// LS Electric XG5000 project: 신호등
// PLC LSPLC

PROGRAM NewProgram (task: 스캔 프로그램)

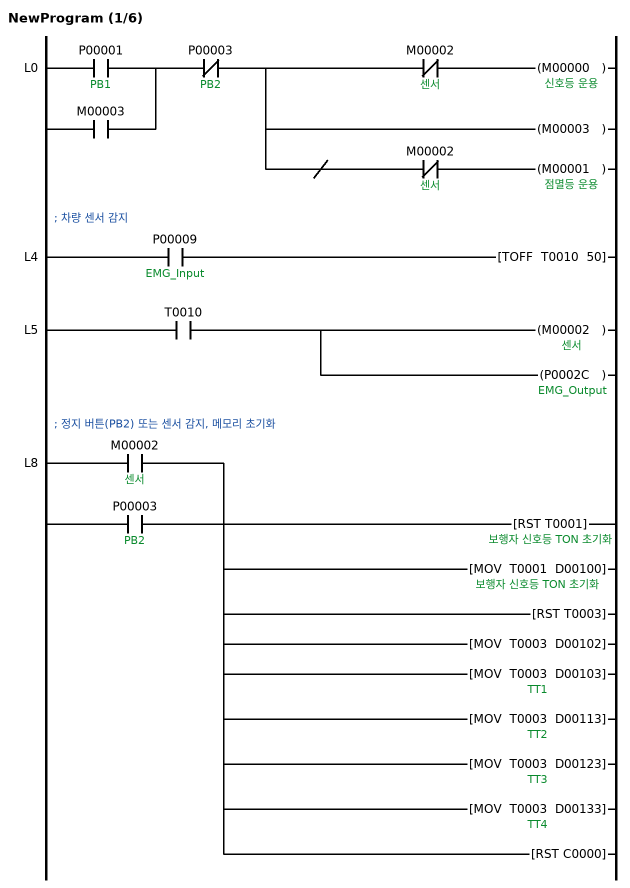
; L0
LOAD      P00001	// PB1
OR        M00003
AND NOT   P00003	// PB2
MPUSH
AND NOT   M00002	// 센서
OUT       M00000	// 신호등 운용
MPOP
OUT       M00003
NOT
AND NOT   M00002	// 센서
OUT       M00001	// 점멸등 운용
// 차량 센서 감지
; L4
LOAD      P00009	// EMG_Input
TOFF      T0010 50
; L5
LOAD      T0010
OUT       M00002	// 센서
OUT       P0002C	// EMG_Output
// 정지 버튼(PB2) 또는 센서 감지, 메모리 초기화
; L8
LOAD      M00002	// 센서
OR        P00003	// PB2
RST       T0001	// 보행자 신호등 TON 초기화
MOV       T0001 D00100	// 보행자 신호등 TON 초기화
RST       T0003
MOV       T0003 D00102
MOV       T0003 D00103	// TT1
MOV       T0003 D00113	// TT2
MOV       T0003 D00123	// TT3
MOV       T0003 D00133	// TT4
RST       C0000

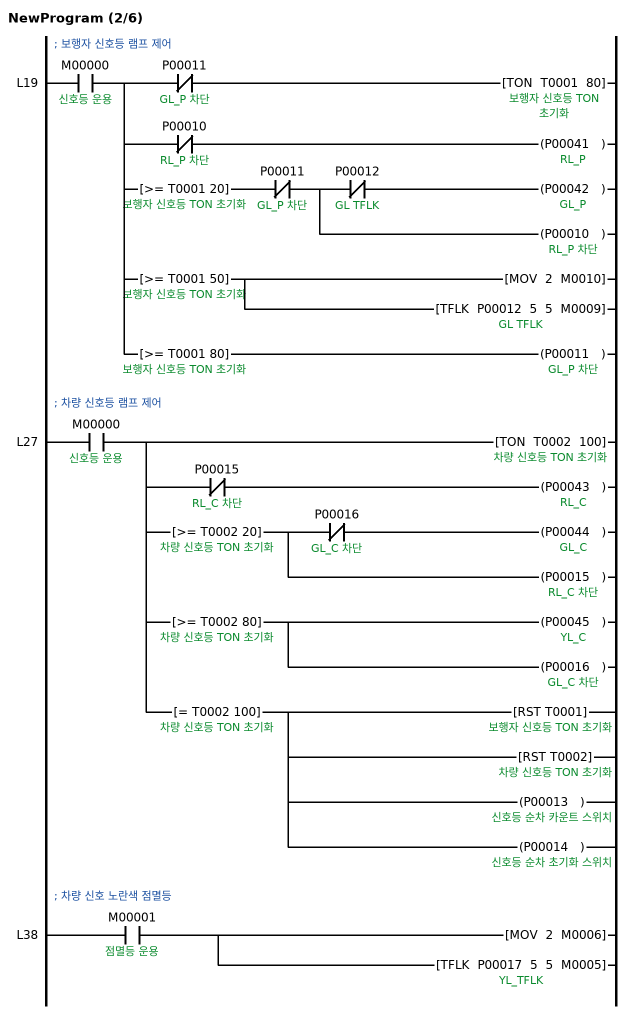
// 보행자 신호등 램프 제어
; L19
LOAD      M00000	// 신호등 운용
MPUSH
AND NOT   P00011	// GL_P 차단
TON       T0001 80	// 보행자 신호등 TON 초기화
MLOAD
AND NOT   P00010	// RL_P 차단
OUT       P00041	// RL_P
MLOAD
AND>=     T0001 20	// 보행자 신호등 TON 초기화
AND NOT   P00011	// GL_P 차단
MPUSH
AND NOT   P00012	// GL TFLK
OUT       P00042	// GL_P
MPOP
OUT       P00010	// RL_P 차단
MLOAD
AND>=     T0001 50	// 보행자 신호등 TON 초기화
MOV       2 M0010
TFLK      P00012 5 5 M0009	// GL TFLK
MPOP
AND>=     T0001 80	// 보행자 신호등 TON 초기화
OUT       P00011	// GL_P 차단
// 차량 신호등 램프 제어
; L27
LOAD      M00000	// 신호등 운용
TON       T0002 100	// 차량 신호등 TON 초기화
MPUSH
AND NOT   P00015	// RL_C 차단
OUT       P00043	// RL_C
MLOAD
AND>=     T0002 20	// 차량 신호등 TON 초기화
MPUSH
AND NOT   P00016	// GL_C 차단
OUT       P00044	// GL_C
MPOP
OUT       P00015	// RL_C 차단
MLOAD
AND>=     T0002 80	// 차량 신호등 TON 초기화
OUT       P00045	// YL_C
OUT       P00016	// GL_C 차단
MPOP
AND=      T0002 100	// 차량 신호등 TON 초기화
RST       T0001	// 보행자 신호등 TON 초기화
RST       T0002	// 차량 신호등 TON 초기화
OUT       P00013	// 신호등 순차 카운트 스위치
OUT       P00014	// 신호등 순차 초기화 스위치
// 차량 신호 노란색 점멸등
; L38
LOAD      M00001	// 점멸등 운용
MOV       2 M0006
TFLK      P00017 5 5 M0005	// YL_TFLK

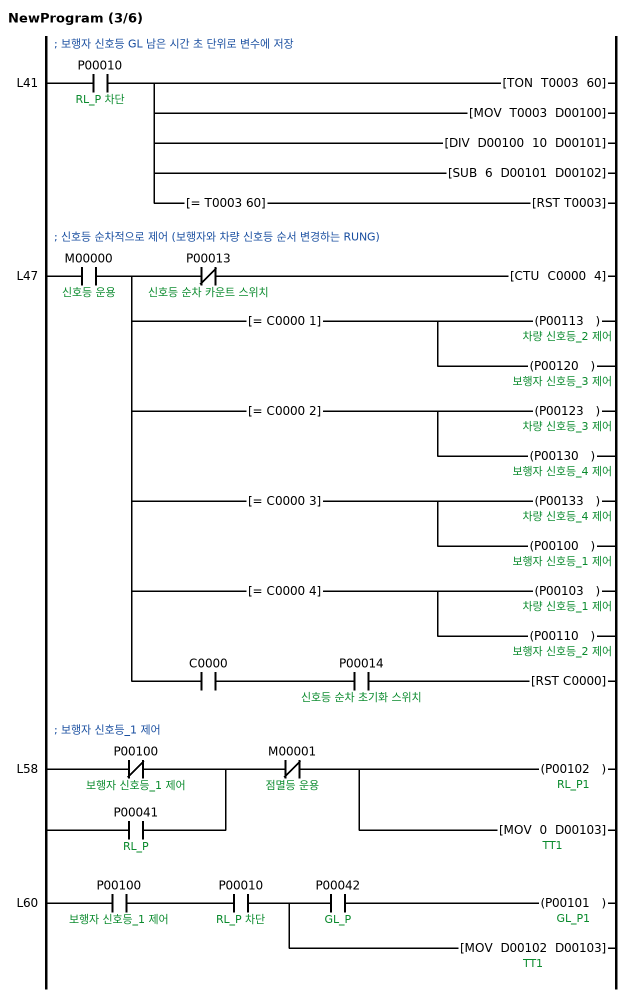
// 보행자 신호등 GL 남은 시간 초 단위로 변수에 저장
; L41
LOAD      P00010	// RL_P 차단
TON       T0003 60
MOV       T0003 D00100
DIV       D00100 10 D00101
SUB       6 D00101 D00102
AND=      T0003 60
RST       T0003
// 신호등 순차적으로 제어 (보행자와 차량 신호등 순서 변경하는 RUNG)
; L47
LOAD      M00000	// 신호등 운용
MPUSH
AND NOT   P00013	// 신호등 순차 카운트 스위치
CTU       C0000 4
MLOAD
AND=      C0000 1
OUT       P00113	// 차량 신호등_2 제어
OUT       P00120	// 보행자 신호등_3 제어
MLOAD
AND=      C0000 2
OUT       P00123	// 차량 신호등_3 제어
OUT       P00130	// 보행자 신호등_4 제어
MLOAD
AND=      C0000 3
OUT       P00133	// 차량 신호등_4 제어
OUT       P00100	// 보행자 신호등_1 제어
MLOAD
AND=      C0000 4
OUT       P00103	// 차량 신호등_1 제어
OUT       P00110	// 보행자 신호등_2 제어
MPOP
AND       C0000
AND       P00014	// 신호등 순차 초기화 스위치
RST       C0000
// 보행자 신호등_1 제어
; L58
LOAD NOT  P00100	// 보행자 신호등_1 제어
OR        P00041	// RL_P
AND NOT   M00001	// 점멸등 운용
OUT       P00102	// RL_P1
MOV       0 D00103	// TT1
; L60
LOAD      P00100	// 보행자 신호등_1 제어
AND       P00010	// RL_P 차단
MPUSH
AND       P00042	// GL_P
OUT       P00101	// GL_P1
MPOP
MOV       D00102 D00103	// TT1

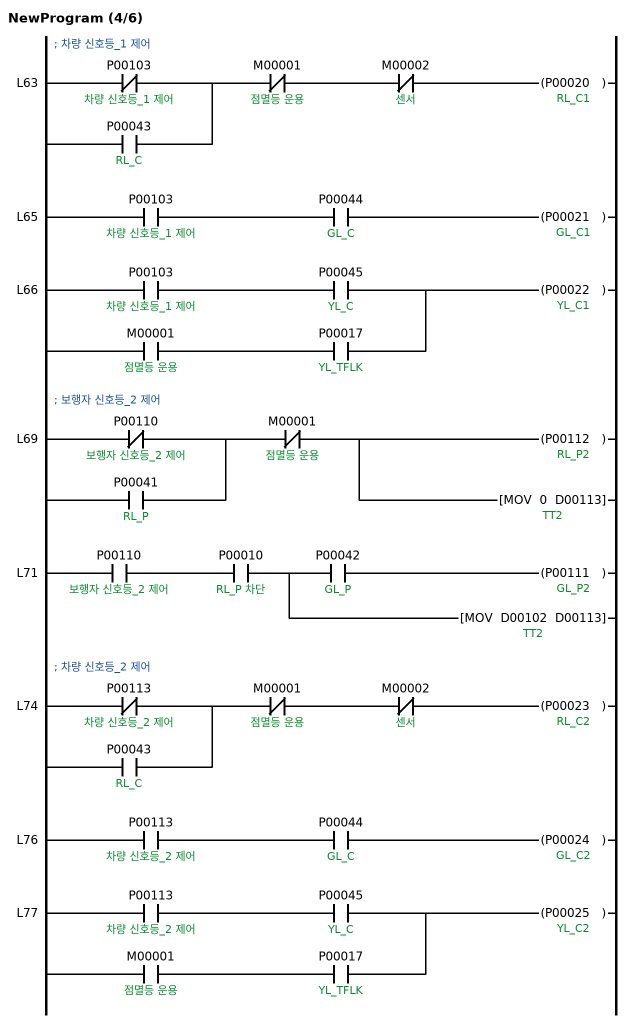
// 차량 신호등_1 제어
; L63
LOAD NOT  P00103	// 차량 신호등_1 제어
OR        P00043	// RL_C
AND NOT   M00001	// 점멸등 운용
AND NOT   M00002	// 센서
OUT       P00020	// RL_C1
; L65
LOAD      P00103	// 차량 신호등_1 제어
AND       P00044	// GL_C
OUT       P00021	// GL_C1
; L66
LOAD      P00103	// 차량 신호등_1 제어
AND       P00045	// YL_C
LOAD      M00001	// 점멸등 운용
AND       P00017	// YL_TFLK
OR LOAD
OUT       P00022	// YL_C1
// 보행자 신호등_2 제어
; L69
LOAD NOT  P00110	// 보행자 신호등_2 제어
OR        P00041	// RL_P
AND NOT   M00001	// 점멸등 운용
OUT       P00112	// RL_P2
MOV       0 D00113	// TT2
; L71
LOAD      P00110	// 보행자 신호등_2 제어
AND       P00010	// RL_P 차단
MPUSH
AND       P00042	// GL_P
OUT       P00111	// GL_P2
MPOP
MOV       D00102 D00113	// TT2
// 차량 신호등_2 제어
; L74
LOAD NOT  P00113	// 차량 신호등_2 제어
OR        P00043	// RL_C
AND NOT   M00001	// 점멸등 운용
AND NOT   M00002	// 센서
OUT       P00023	// RL_C2
; L76
LOAD      P00113	// 차량 신호등_2 제어
AND       P00044	// GL_C
OUT       P00024	// GL_C2
; L77
LOAD      P00113	// 차량 신호등_2 제어
AND       P00045	// YL_C
LOAD      M00001	// 점멸등 운용
AND       P00017	// YL_TFLK
OR LOAD
OUT       P00025	// YL_C2

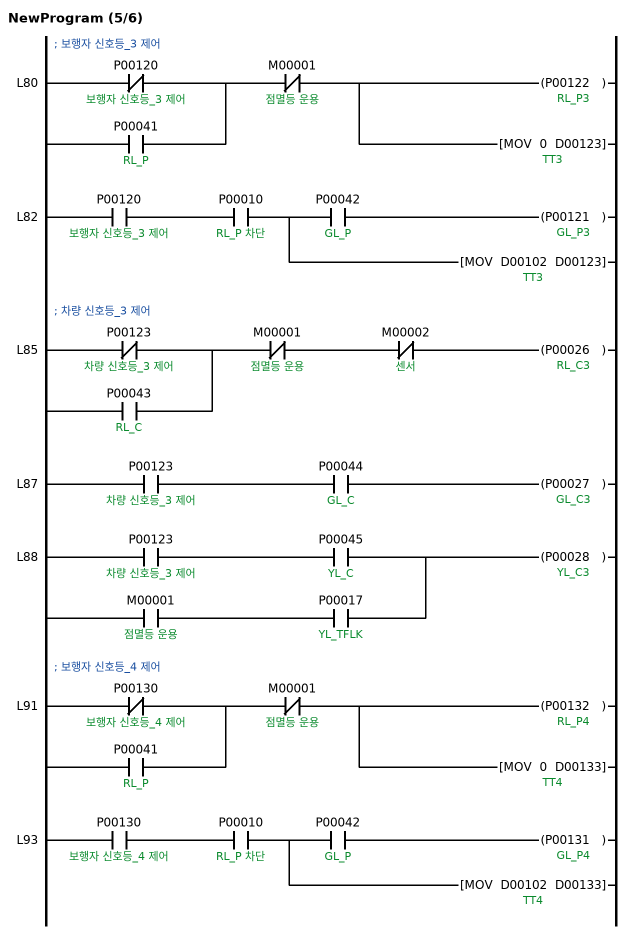
// 보행자 신호등_3 제어
; L80
LOAD NOT  P00120	// 보행자 신호등_3 제어
OR        P00041	// RL_P
AND NOT   M00001	// 점멸등 운용
OUT       P00122	// RL_P3
MOV       0 D00123	// TT3
; L82
LOAD      P00120	// 보행자 신호등_3 제어
AND       P00010	// RL_P 차단
MPUSH
AND       P00042	// GL_P
OUT       P00121	// GL_P3
MPOP
MOV       D00102 D00123	// TT3
// 차량 신호등_3 제어
; L85
LOAD NOT  P00123	// 차량 신호등_3 제어
OR        P00043	// RL_C
AND NOT   M00001	// 점멸등 운용
AND NOT   M00002	// 센서
OUT       P00026	// RL_C3
; L87
LOAD      P00123	// 차량 신호등_3 제어
AND       P00044	// GL_C
OUT       P00027	// GL_C3
; L88
LOAD      P00123	// 차량 신호등_3 제어
AND       P00045	// YL_C
LOAD      M00001	// 점멸등 운용
AND       P00017	// YL_TFLK
OR LOAD
OUT       P00028	// YL_C3
// 보행자 신호등_4 제어
; L91
LOAD NOT  P00130	// 보행자 신호등_4 제어
OR        P00041	// RL_P
AND NOT   M00001	// 점멸등 운용
OUT       P00132	// RL_P4
MOV       0 D00133	// TT4
; L93
LOAD      P00130	// 보행자 신호등_4 제어
AND       P00010	// RL_P 차단
MPUSH
AND       P00042	// GL_P
OUT       P00131	// GL_P4
MPOP
MOV       D00102 D00133	// TT4

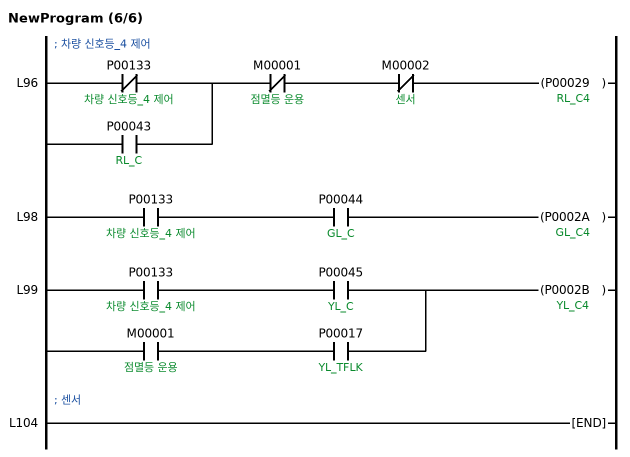
// 차량 신호등_4 제어
; L96
LOAD NOT  P00133	// 차량 신호등_4 제어
OR        P00043	// RL_C
AND NOT   M00001	// 점멸등 운용
AND NOT   M00002	// 센서
OUT       P00029	// RL_C4
; L98
LOAD      P00133	// 차량 신호등_4 제어
AND       P00044	// GL_C
OUT       P0002A	// GL_C4
; L99
LOAD      P00133	// 차량 신호등_4 제어
AND       P00045	// YL_C
LOAD      M00001	// 점멸등 운용
AND       P00017	// YL_TFLK
OR LOAD
OUT       P0002B	// YL_C4
// 센서
; L104
END

VARIABLES AND COMMENTS (devices not used above)
P00004	BIT	PB4